Fanuc KAREL source: KT00904.KL

PROGRAM KT00904
%NOLOCKGROUP
%ENVIRONMENT VECTR
VAR
  P1: XYZWPR
  P2: XYZWPR
  OUT: VECTOR
BEGIN
  P1.X = 1.0
  P2.Y = 2.0
  P1.X = 1.0
  P2.Y = 2.0
  OUT = APPROACH(P1)
END KT00904
